// TIA Portal V20 export
// export: Created 2026-10-12T05:42:34.7676686Z, ExportSetting WithDefaults, DisplayName Totally Integrated Automation Portal, DisplayVersion V20, DisplayName TIA Portal Openness, DisplayVersion V20, DisplayName TIA Portal Teamcenter Gateway, DisplayVersion V20, DisplayName TIA Portal Version Control Interface, DisplayVersion V20, DisplayName SINAMICS Startdrive Advanced, DisplayVersion V20 SP1 Update 2, DisplayName SINAMICS Startdrive G110M, G120, G120C, G120D, G120P, G115D, DisplayVersion V20 SP1 Update 2, DisplayName SINAMICS Startdrive G130, G150, S120, S150, SINAMICS MV, G220, S200, S210, DisplayVersion V20 SP1 Update 2, DisplayName STEP 7 Professional, DisplayVersion V20, DisplayName STEP 7 Safety, DisplayVersion V20, DisplayName WinCC Basic/Comfort/Advanced, DisplayVersion V20, DisplayName WinCC Professional, DisplayVersion V20, DisplayName WinCC Unified, DisplayVersion V20
FUNCTION_BLOCK "FB_PressDemoHome"   // FB4, SCL
{ S7_Optimized_Access := 'TRUE' }
VERSION : 0.1
// stored: AutoNumber true, IsIECCheckEnabled false, IsRetainMemResEnabled false, MemoryReserve 100, SetENOAutomatically false, UDAEnableTagReadback false
   VAR_INPUT
      Run : Bool;
      Reset : Bool;
      OwnerIndex : DInt;
      Delta : Time;
   END_VAR
   VAR_IN_OUT
      PressRam : "FB_CylinderCM";
      Door : "FB_CylinderCM";
      PartSlide : "FB_CylinderCM";
   END_VAR
   VAR
      Seq { ExternalWritable := 'False'; S7_SetPoint := 'True'} : "FRK_SequenceCtx";
      Row1 { ExternalWritable := 'False'; S7_SetPoint := 'True'} : "FRK_SequenceRow";
      Row2 { ExternalWritable := 'False'; S7_SetPoint := 'True'} : "FRK_SequenceRow";
      Row3 { ExternalWritable := 'False'; S7_SetPoint := 'True'} : "FRK_SequenceRow";
      Row4 { ExternalWritable := 'False'; S7_SetPoint := 'True'} : "FRK_SequenceRow";
      At0 { ExternalAccessible := 'False'; ExternalVisible := 'False'; ExternalWritable := 'False'} : Bool;
      At900 { ExternalAccessible := 'False'; ExternalVisible := 'False'; ExternalWritable := 'False'} : Bool;
      At910 { ExternalAccessible := 'False'; ExternalVisible := 'False'; ExternalWritable := 'False'} : Bool;
      At999 { ExternalAccessible := 'False'; ExternalVisible := 'False'; ExternalWritable := 'False'} : Bool;
      Ready1 { ExternalAccessible := 'False'; ExternalVisible := 'False'; ExternalWritable := 'False'} : Bool;
      Ready2 { ExternalAccessible := 'False'; ExternalVisible := 'False'; ExternalWritable := 'False'} : Bool;
      Ready3 { ExternalAccessible := 'False'; ExternalVisible := 'False'; ExternalWritable := 'False'} : Bool;
      Ready4 { ExternalAccessible := 'False'; ExternalVisible := 'False'; ExternalWritable := 'False'} : Bool;
      Ready5 { ExternalAccessible := 'False'; ExternalVisible := 'False'; ExternalWritable := 'False'} : Bool;
      Advance { ExternalAccessible := 'False'; ExternalVisible := 'False'; ExternalWritable := 'False'} : Bool;
   END_VAR
BEGIN

   "FRK_SeqBegin"(Run := #Run,
                  Reset := #Reset,
                  OwnerIndex := #OwnerIndex,
                  ChainIndex := 2,
                  BranchIndex := 0,
                  Delta := #Delta,
                  Seq := #Seq);
   "F_CylinderSequenceLease"(Seq := #Seq,
                             Target := #PressRam);
   "F_CylinderSequenceLease"(Seq := #Seq,
                             Target := #Door);
   "F_CylinderSequenceLease"(Seq := #Seq,
                             Target := #PartSlide);
   CASE #Seq.ScanStep OF
       0:
           IF #Seq.Running AND NOT #Seq.Error THEN
               "FRK_SeqStep"(StepNo := 0,
                             StepName := 'project.step.pressHomeInitialize',
                             Seq := #Seq,
                             Row := #Row1);
               "FRK_SeqReady"(Seq := #Seq,
                              Ok1 := TRUE,
                              Ok2 := TRUE,
                              Ok3 := TRUE,
                              Ok4 := TRUE,
                              Ok5 := TRUE);
               "FRK_SeqRoute"(Seq := #Seq,
                              OnAdvance := 900,
                              OnJump1 := -1);
           END_IF;
       900:
           IF #Seq.Running AND NOT #Seq.Error THEN
               "FRK_SeqStep"(StepNo := 900,
                             StepName := 'project.step.pressHomeRam',
                             Seq := #Seq,
                             Row := #Row2);
               #Ready1 := "F_CylinderRetract"(Seq := #Seq, Target := #PressRam);
               "FRK_SeqReady"(Seq := #Seq,
                              Ok1 := #Ready1,
                              Ok2 := TRUE,
                              Ok3 := TRUE,
                              Ok4 := TRUE,
                              Ok5 := TRUE);
               "FRK_SeqRoute"(Seq := #Seq,
                              OnAdvance := 910,
                              OnJump1 := -1);
           END_IF;
       910:
           IF #Seq.Running AND NOT #Seq.Error THEN
               "FRK_SeqStep"(StepNo := 910,
                             StepName := 'project.step.pressHomeDoorAndSlide',
                             Seq := #Seq,
                             Row := #Row3);
               #Ready1 := "F_CylinderRetract"(Seq := #Seq, Target := #Door);
               #Ready2 := "F_CylinderRetract"(Seq := #Seq, Target := #PartSlide);
               "FRK_SeqReady"(Seq := #Seq,
                              Ok1 := #Ready1,
                              Ok2 := #Ready2,
                              Ok3 := TRUE,
                              Ok4 := TRUE,
                              Ok5 := TRUE);
               "FRK_SeqRoute"(Seq := #Seq,
                              OnAdvance := 999,
                              OnJump1 := -1);
           END_IF;
       999:
           IF #Seq.Running AND NOT #Seq.Error THEN
               "FRK_SeqStep"(StepNo := 999,
                             StepName := 'project.step.pressHomeComplete',
                             Seq := #Seq,
                             Row := #Row4);
               "FRK_SeqComplete"(Seq := #Seq);
           END_IF;
       ELSE
           #Seq.Error := TRUE;
           #Seq.ErrorDiagnostic.ReasonCode := 10001;
           #Seq.ErrorDiagnostic.Description := WSTRING#'project.sequence.invalidStep';
   END_CASE;
   "F_CylinderSequenceLease"(Seq := #Seq,
                             Target := #PressRam);
   "F_CylinderSequenceLease"(Seq := #Seq,
                             Target := #Door);
   "F_CylinderSequenceLease"(Seq := #Seq,
                             Target := #PartSlide);
END_FUNCTION_BLOCK
